TYPE ST_EL3312CoeWriteData_1 :
STRUCT
	wIdx: WORD;
	bySubIdx: BYTE;
	bWriteOK: BOOL;
	dwData: DWORD;
	nSize: UDINT;
END_STRUCT
END_TYPE

(* stored: Version 1.1.0.1, ProductVersion 3.1.4024.15
   DUT ST_EL3312CoeWriteData_1: Id {cea9fb03-f4e9-48c7-b924-631091eda557} *)
